METHOD PUBLIC Cyclic
VAR_INPUT
    eMode                    : E_PuckLockerMode;
    bSensorUp                : BOOL;
    bSensorDown              : BOOL;
    bPartRemovedFromNest     : BOOL;
    bReleasePassPuck         : BOOL;
    bAcknowledgeFault        : BOOL;
    bEmptyPuckBypass         : BOOL;
    tRemovalConfirm          : TIME;
END_VAR
VAR_OUTPUT bPinCommandUp : BOOL; END_VAR
bEnabledInternal := eMode <> E_PuckLockerMode.Disabled;
bDetectedInternal := bSensorUp OR bSensorDown;
bAckPulseInternal := bAcknowledgeFault AND NOT bAcknowledgePrevious;
bAcknowledgePrevious := bAcknowledgeFault;

stStatusInternal.eMode := eMode;
stStatusInternal.bPuckDetected := bDetectedInternal;
stStatusInternal.bPuckSensorMismatch := bSensorUp XOR bSensorDown;
stStatusInternal.bPuckLocked := bPinCommandUp AND bDetectedInternal;
stStatusInternal.bMachinePermissive := NOT stStatusInternal.bUnexpectedRemovalFault AND NOT stStatusInternal.bPuckSensorMismatch;
stStatusInternal.bIndexPermissive := stStatusInternal.bMachinePermissive AND eState <> E_PuckLockerState.UnexpectedPuckRemovalFault;

IF bReleasePassPuck THEN bReleaseRequested := TRUE; END_IF
IF bPartRemovedFromNest THEN bPartRemoved := TRUE; END_IF

CASE eState OF
E_PuckLockerState.Disabled:
    bPinCommandUp := FALSE;
    stStatusInternal.bRemovalAllowed := TRUE;
    stStatusInternal.sMessage := 'Puck locker disabled';
    bReleaseRequested := FALSE; bPartRemoved := FALSE;
    IF bEnabledInternal THEN
        IF bDetectedInternal THEN eState := E_PuckLockerState.LockingPuck; ELSE eState := E_PuckLockerState.WaitingForPuck; END_IF
    END_IF

E_PuckLockerState.WaitingForPuck:
    bPinCommandUp := FALSE;
    stStatusInternal.bRemovalAllowed := TRUE;
    stStatusInternal.sMessage := 'Load puck';
    IF NOT bEnabledInternal THEN eState := E_PuckLockerState.Disabled;
    ELSIF bDetectedInternal THEN eState := E_PuckLockerState.LockingPuck;
    END_IF

E_PuckLockerState.LockingPuck:
    bPinCommandUp := TRUE;
    stStatusInternal.bRemovalAllowed := FALSE;
    stStatusInternal.sMessage := 'Locking puck';
    IF NOT bEnabledInternal THEN eState := E_PuckLockerState.Disabled;
    ELSIF bDetectedInternal THEN eState := E_PuckLockerState.Locked;
    END_IF

E_PuckLockerState.Locked:
    bPinCommandUp := TRUE;
    stStatusInternal.bRemovalAllowed := FALSE;
    stStatusInternal.sMessage := 'Puck locked';
    IF NOT bEnabledInternal THEN eState := E_PuckLockerState.Disabled;
    ELSIF NOT bDetectedInternal THEN
        stStatusInternal.bUnexpectedRemovalFault := TRUE;
        eState := E_PuckLockerState.UnexpectedPuckRemovalFault;
    ELSIF bReleaseRequested THEN
        eState := E_PuckLockerState.WaitingForPartRemoval;
    ELSIF bEmptyPuckBypass AND eMode = E_PuckLockerMode.EnabledWithEmptyPuckBypass THEN
        eState := E_PuckLockerState.ReleasingPuck;
    END_IF

E_PuckLockerState.WaitingForPartRemoval:
    bPinCommandUp := TRUE;
    stStatusInternal.sMessage := 'Remove processed part';
    IF NOT bDetectedInternal THEN
        stStatusInternal.bUnexpectedRemovalFault := TRUE;
        eState := E_PuckLockerState.UnexpectedPuckRemovalFault;
    ELSIF bPartRemoved THEN eState := E_PuckLockerState.ReleasingPuck;
    END_IF

E_PuckLockerState.ReleasingPuck:
    bPinCommandUp := FALSE;
    stStatusInternal.bRemovalAllowed := TRUE;
    stStatusInternal.sMessage := 'Remove released puck';
    tonRemovalConfirm(IN := NOT bDetectedInternal, PT := tRemovalConfirm);
    IF tonRemovalConfirm.Q THEN
        bReleaseRequested := FALSE; bPartRemoved := FALSE;
        tonRemovalConfirm(IN := FALSE);
        eState := E_PuckLockerState.WaitingForPuck;
    END_IF

E_PuckLockerState.UnexpectedPuckRemovalFault:
    bPinCommandUp := TRUE;
    stStatusInternal.bUnexpectedRemovalFault := TRUE;
    stStatusInternal.sMessage := 'Restore puck and acknowledge';
    IF bAckPulseInternal AND bDetectedInternal THEN
        stStatusInternal.bUnexpectedRemovalFault := FALSE;
        eState := E_PuckLockerState.Locked;
    END_IF
END_CASE

stStatusInternal.eState := eState;
stStatusInternal.bReleaseRequested := bReleaseRequested;
stStatusInternal.bPartRemovalConfirmed := bPartRemoved;
stStatusInternal.bDispositionPending := bReleaseRequested OR (eState = E_PuckLockerState.WaitingForPartRemoval) OR (eState = E_PuckLockerState.ReleasingPuck);
stStatusInternal.bPuckLocked := bPinCommandUp AND bDetectedInternal;
stStatusInternal.bIndexPermissive := NOT stStatusInternal.bUnexpectedRemovalFault AND NOT stStatusInternal.bPuckSensorMismatch;
stStatusInternal.bMachinePermissive := stStatusInternal.bIndexPermissive;
bPreviousPuckDetected := bDetectedInternal;
END_METHOD

METHOD PUBLIC GetStatus : ST_PuckLockerStatus
GetStatus := stStatusInternal;
END_METHOD

METHOD PUBLIC IsFaulted : BOOL
IsFaulted := stStatusInternal.bUnexpectedRemovalFault OR stStatusInternal.bPuckSensorMismatch;
END_METHOD

METHOD PUBLIC IsLocked : BOOL
IsLocked := stStatusInternal.bPuckLocked AND eState = E_PuckLockerState.Locked;
END_METHOD

END_FUNCTION_BLOCK

// ---- POUs/02_Components/Pneumatics/FB_Support.TcPOU
FUNCTION_BLOCK FB_Support
VAR
    tonMovementTimeout : TON;

    bFaultInternal     : BOOL;
    bExtendOutputInternal  : BOOL;
    bRetractOutputInternal : BOOL;
END_VAR

METHOD PUBLIC Cyclic
VAR_INPUT
    bEnable          : BOOL;
    bRaiseRequest    : BOOL;
    bLowerRequest    : BOOL;
    bStopRequest     : BOOL;

    bExtended        : BOOL;
    bRetracted       : BOOL;

    tMovementTimeout : TIME;
END_VAR

VAR_OUTPUT
    bExtendOutput    : BOOL;
    bRetractOutput   : BOOL;
END_VAR
// =========================================================
// DEFAULT OUTPUTS
// =========================================================

bExtendOutputInternal := FALSE;
bRetractOutputInternal := FALSE;


// =========================================================
// FAULT DETECTION
// =========================================================

IF bExtended AND bRetracted THEN
    bFaultInternal := TRUE;
END_IF

IF bRaiseRequest AND bLowerRequest THEN
    bFaultInternal := TRUE;
END_IF


// =========================================================
// STOP HANDLING
// =========================================================
//
// Stop does not reset the component.
// Stop commands the station support to its safe position.

IF bStopRequest THEN

    tonMovementTimeout(
        IN := NOT bRetracted,
        PT := tMovementTimeout
    );

    IF NOT bRetracted AND NOT bFaultInternal THEN
        bRetractOutputInternal := TRUE;
    END_IF

    IF tonMovementTimeout.Q THEN
        bFaultInternal := TRUE;
    END_IF


// =========================================================
// COMPONENT DISABLED OR FAULTED
// =========================================================

ELSIF NOT bEnable OR bFaultInternal THEN

    tonMovementTimeout(IN := FALSE);


// =========================================================
// NORMAL MOVEMENT CONTROL
// =========================================================

ELSE

    // -----------------------------------------------------
    // EXTEND
    // -----------------------------------------------------

    IF bRaiseRequest AND NOT bLowerRequest THEN

        tonMovementTimeout(
            IN := (GVL_MASTER.stStatus.eMachineState <> E_MachineState.Manual)
        AND NOT bExtended, 
            PT := tMovementTimeout
        );

        IF NOT bExtended THEN
            bExtendOutputInternal := TRUE;
        END_IF

        IF tonMovementTimeout.Q THEN
            bFaultInternal := TRUE;
        END_IF


    // -----------------------------------------------------
    // RETRACT
    // -----------------------------------------------------

    ELSIF bLowerRequest AND NOT bRaiseRequest THEN

        tonMovementTimeout(
            IN := (GVL_MASTER.stStatus.eMachineState <> E_MachineState.Manual)
        AND NOT bRetracted,
            PT := tMovementTimeout
        );

        IF NOT bRetracted THEN
            bRetractOutputInternal := TRUE;
        END_IF

        IF tonMovementTimeout.Q THEN
            bFaultInternal := TRUE;
        END_IF


    // -----------------------------------------------------
    // NO COMMAND
    // -----------------------------------------------------

    ELSE

        tonMovementTimeout(IN := FALSE);

    END_IF

END_IF


// =========================================================
// OUTPUT MAPPING
// =========================================================

bExtendOutput := bExtendOutputInternal;
bRetractOutput := bRetractOutputInternal;
END_METHOD

METHOD IsFaulted : BOOL
VAR_INPUT
END_VAR
IsFaulted := bFaultInternal;
END_METHOD

METHOD PUBLIC Reset
bFaultInternal := FALSE;

bExtendOutputInternal := FALSE;
bRetractOutputInternal := FALSE;

tonMovementTimeout(IN := FALSE);
END_METHOD

END_FUNCTION_BLOCK

// ---- POUs/06_Utilities/F_ScaleLinear.TcPOU
FUNCTION F_ScaleLinear : REAL
VAR_INPUT
    rRawValue : REAL;
    rRawMin   : REAL;
    rRawMax   : REAL;
    rEngMin   : REAL;
    rEngMax   : REAL;
END_VAR
VAR
    rSpanRaw : REAL;
END_VAR

rSpanRaw := rRawMax - rRawMin;

IF ABS(rSpanRaw) > 0.000001 THEN

    F_ScaleLinear :=
        ((rRawValue - rRawMin) / rSpanRaw)
        * (rEngMax - rEngMin)
        + rEngMin;

ELSE

    F_ScaleLinear := rEngMin;

END_IF

END_FUNCTION
